(* IEC 61131-3 sources: PLC-Static-Analysis/modules/plc-rules/src/test/resources/PLCA-L018, 2 files *)

(* ---- compliant.st ---- *)
PROGRAM P_L018ok
VAR
    n : INT;
    m : INT;
    r : REAL;
    b : BOOL;
    c : BOOL;
    q : BOOL;
END_VAR
IF n < 10 THEN
    ; // nothing below the limit: the pump keeps its state
ELSE
    q := TRUE;
END_IF
IF n >= 10 THEN
    q := TRUE;
END_IF
END_PROGRAM

(* ---- noncompliant.st ---- *)
PROGRAM P_L018
VAR
    n : INT;
    m : INT;
    r : REAL;
    b : BOOL;
    c : BOOL;
    q : BOOL;
END_VAR
(* PLCA-L018 *) IF n < 10 THEN
ELSE
    q := TRUE;
END_IF
END_PROGRAM
